Fanuc KAREL source: kb00168.KL

-- PROVISIONAL review KL for V770-1; original PC SHA256 2c69c0a73fad8c839bfb57f40c3790f0c382114ea0e20c6ff051d336708c2b48
-- Incomplete behavior may be omitted. Consult companion uncertainty JSON. Do not deploy.
PROGRAM KB00168
%NOLOCKGROUP
BEGIN
  -- UNRESOLVED_PC offsets 5-14; opcodes 3F,75
  -- UNRESOLVED_PC offsets 19-26; opcodes 9D,23
  -- UNRESOLVED_PC offsets 31-49; opcodes 27,22,2A,22,31
  -- UNRESOLVED_PC offsets 54-58; opcodes 7F
END KB00168
